(* IEC 61131-3 sources: daoli-st-library/_tools/rusty, 1 file *)

(* ---- iec_std_stub.st ---- *)
(* ============================================================================
   iec_std_stub.st  ——  道莅 L2 编译闸：IEC 61131-3 标准库外部声明桩
   ----------------------------------------------------------------------------
   用途：RuSTy (plc.exe) 不内建 IEC 标准函数/标准 FB 的声明，裸编译会把
        ABS/TON/R_TRIG 等判为 "Unknown type / Could not resolve reference"。
        本文件以 {external} 声明标准件接口，仅作 --check 夹具，不产生实现。

   纪律：
   1. 本文件**不属于**代码库交付物，只放在 _tools/rusty/ 下，不入 INDEX_REGISTRY。
   2. 声明按 IEC 61131-3 第 3 版标准语义书写，与各件源码零耦合。
   3. 泛型用 ANY_NUM / ANY_ELEMENTARY 表达，避免为每种位宽写重复声明。
   ============================================================================ *)

{external}
FUNCTION ABS<T: ANY_NUM> : T
VAR_INPUT IN : T; END_VAR
END_FUNCTION

{external}
FUNCTION SQRT<T: ANY_REAL> : T
VAR_INPUT IN : T; END_VAR
END_FUNCTION

{external}
FUNCTION LN<T: ANY_REAL> : T
VAR_INPUT IN : T; END_VAR
END_FUNCTION

{external}
FUNCTION LOG<T: ANY_REAL> : T
VAR_INPUT IN : T; END_VAR
END_FUNCTION

{external}
FUNCTION EXP<T: ANY_REAL> : T
VAR_INPUT IN : T; END_VAR
END_FUNCTION

{external}
FUNCTION SIN<T: ANY_REAL> : T
VAR_INPUT IN : T; END_VAR
END_FUNCTION

{external}
FUNCTION COS<T: ANY_REAL> : T
VAR_INPUT IN : T; END_VAR
END_FUNCTION

{external}
FUNCTION TAN<T: ANY_REAL> : T
VAR_INPUT IN : T; END_VAR
END_FUNCTION

{external}
FUNCTION ASIN<T: ANY_REAL> : T
VAR_INPUT IN : T; END_VAR
END_FUNCTION

{external}
FUNCTION ACOS<T: ANY_REAL> : T
VAR_INPUT IN : T; END_VAR
END_FUNCTION

{external}
FUNCTION ATAN<T: ANY_REAL> : T
VAR_INPUT IN : T; END_VAR
END_FUNCTION

{external}
FUNCTION EXPT<T: ANY_REAL> : T
VAR_INPUT IN1 : T; IN2 : T; END_VAR
END_FUNCTION

{external}
FUNCTION TRUNC<T: ANY_REAL> : T
VAR_INPUT IN : T; END_VAR
END_FUNCTION

{external}
FUNCTION ROUND<T: ANY_REAL> : T
VAR_INPUT IN : T; END_VAR
END_FUNCTION

{external}
FUNCTION FLOOR<T: ANY_REAL> : T
VAR_INPUT IN : T; END_VAR
END_FUNCTION

{external}
FUNCTION CEIL<T: ANY_REAL> : T
VAR_INPUT IN : T; END_VAR
END_FUNCTION

{external}
FUNCTION MIN<T: ANY_ELEMENTARY> : T
VAR_INPUT IN1 : T; IN2 : T; END_VAR
END_FUNCTION

{external}
FUNCTION MAX<T: ANY_ELEMENTARY> : T
VAR_INPUT IN1 : T; IN2 : T; END_VAR
END_FUNCTION

{external}
FUNCTION LIMIT<T: ANY_ELEMENTARY> : T
VAR_INPUT MN : T; IN : T; MX : T; END_VAR
END_FUNCTION

{external}
FUNCTION SEL<T: ANY_ELEMENTARY> : T
VAR_INPUT G : BOOL; IN0 : T; IN1 : T; END_VAR
END_FUNCTION

{external}
FUNCTION MUX<T: ANY_ELEMENTARY> : T
VAR_INPUT K : INT; IN0 : T; IN1 : T; IN2 : T; IN3 : T; END_VAR
END_FUNCTION

{external}
FUNCTION SHL<T: ANY_BIT> : T
VAR_INPUT IN : T; N : INT; END_VAR
END_FUNCTION

{external}
FUNCTION SHR<T: ANY_BIT> : T
VAR_INPUT IN : T; N : INT; END_VAR
END_FUNCTION

{external}
FUNCTION ROL<T: ANY_BIT> : T
VAR_INPUT IN : T; N : INT; END_VAR
END_FUNCTION

{external}
FUNCTION ROR<T: ANY_BIT> : T
VAR_INPUT IN : T; N : INT; END_VAR
END_FUNCTION

(* ---- 字符串九函数 ---- *)
{external}
FUNCTION LEN : UDINT
VAR_INPUT IN : STRING; END_VAR
END_FUNCTION

{external}
FUNCTION LEFT : STRING
VAR_INPUT IN : STRING; L : UDINT; END_VAR
END_FUNCTION

{external}
FUNCTION RIGHT : STRING
VAR_INPUT IN : STRING; L : UDINT; END_VAR
END_FUNCTION

{external}
FUNCTION MID : STRING
VAR_INPUT IN : STRING; L : UDINT; P : UDINT := 1; END_VAR
END_FUNCTION

{external}
FUNCTION CONCAT : STRING
VAR_INPUT IN1 : STRING; IN2 : STRING := ''; IN3 : STRING := ''; IN4 : STRING := ''; END_VAR
END_FUNCTION

{external}
FUNCTION INSERT : STRING
VAR_INPUT IN1 : STRING; IN2 : STRING; P : UDINT; END_VAR
END_FUNCTION

{external}
FUNCTION DELETE : STRING
VAR_INPUT IN : STRING; L : UDINT; P : UDINT; END_VAR
END_FUNCTION

{external}
FUNCTION REPLACE : STRING
VAR_INPUT IN1 : STRING; IN2 : STRING; L : UDINT; P : UDINT; END_VAR
END_FUNCTION

{external}
FUNCTION FIND : UDINT
VAR_INPUT IN1 : STRING; IN2 : STRING; END_VAR
END_FUNCTION

{external}
FUNCTION STRING_EQUAL : BOOL
VAR_INPUT a : STRING; b : STRING; END_VAR
END_FUNCTION

{external}
FUNCTION STRING_GREATER : BOOL
VAR_INPUT a : STRING; b : STRING; END_VAR
END_FUNCTION

{external}
FUNCTION STRING_LESS : BOOL
VAR_INPUT a : STRING; b : STRING; END_VAR
END_FUNCTION

{external}
FUNCTION WSTRING_EQUAL : BOOL
VAR_INPUT a : WSTRING; b : WSTRING; END_VAR
END_FUNCTION

(* ---- 标准边沿/定时/计数 FB（空体声明，仅满足类型解析） ---- *)
FUNCTION_BLOCK TON
VAR_INPUT
    IN : BOOL;
    PT : TIME;
END_VAR
VAR_OUTPUT
    Q : BOOL;
    ET : TIME;
END_VAR
END_FUNCTION_BLOCK

FUNCTION_BLOCK TOF
VAR_INPUT
    IN : BOOL;
    PT : TIME;
END_VAR
VAR_OUTPUT
    Q : BOOL;
    ET : TIME;
END_VAR
END_FUNCTION_BLOCK

FUNCTION_BLOCK TP
VAR_INPUT
    IN : BOOL;
    PT : TIME;
END_VAR
VAR_OUTPUT
    Q : BOOL;
    ET : TIME;
END_VAR
END_FUNCTION_BLOCK

FUNCTION_BLOCK R_TRIG
VAR_INPUT
    CLK : BOOL;
END_VAR
VAR_OUTPUT
    Q : BOOL;
END_VAR
END_FUNCTION_BLOCK

FUNCTION_BLOCK F_TRIG
VAR_INPUT
    CLK : BOOL;
END_VAR
VAR_OUTPUT
    Q : BOOL;
END_VAR
END_FUNCTION_BLOCK

FUNCTION_BLOCK CTU
VAR_INPUT
    CU : BOOL;
    R : BOOL;
    PV : INT;
END_VAR
VAR_OUTPUT
    Q : BOOL;
    CV : INT;
END_VAR
END_FUNCTION_BLOCK

FUNCTION_BLOCK CTD
VAR_INPUT
    CD : BOOL;
    LD : BOOL;
    PV : INT;
END_VAR
VAR_OUTPUT
    Q : BOOL;
    CV : INT;
END_VAR
END_FUNCTION_BLOCK

FUNCTION_BLOCK CTUD
VAR_INPUT
    CU : BOOL;
    CD : BOOL;
    R : BOOL;
    LD : BOOL;
    PV : INT;
END_VAR
VAR_OUTPUT
    QU : BOOL;
    QD : BOOL;
    CV : INT;
END_VAR
END_FUNCTION_BLOCK

(* ---- R71 补：类型转换 / ATAN2 / MOVE ---- *)
{external}
FUNCTION TIME_TO_REAL : REAL
VAR_INPUT IN : TIME; END_VAR
END_FUNCTION

{external}
FUNCTION TIME_TO_LREAL : LREAL
VAR_INPUT IN : TIME; END_VAR
END_FUNCTION

{external}
FUNCTION TIME_TO_DINT : DINT
VAR_INPUT IN : TIME; END_VAR
END_FUNCTION

{external}
FUNCTION TIME_TO_UDINT : UDINT
VAR_INPUT IN : TIME; END_VAR
END_FUNCTION

{external}
FUNCTION TIME_TO_LINT : LINT
VAR_INPUT IN : TIME; END_VAR
END_FUNCTION

{external}
FUNCTION UDINT_TO_REAL : REAL
VAR_INPUT IN : UDINT; END_VAR
END_FUNCTION

{external}
FUNCTION UDINT_TO_LREAL : LREAL
VAR_INPUT IN : UDINT; END_VAR
END_FUNCTION

{external}
FUNCTION UDINT_TO_DINT : DINT
VAR_INPUT IN : UDINT; END_VAR
END_FUNCTION

{external}
FUNCTION DINT_TO_REAL : REAL
VAR_INPUT IN : DINT; END_VAR
END_FUNCTION

{external}
FUNCTION DINT_TO_LREAL : LREAL
VAR_INPUT IN : DINT; END_VAR
END_FUNCTION

{external}
FUNCTION INT_TO_REAL : REAL
VAR_INPUT IN : INT; END_VAR
END_FUNCTION

{external}
FUNCTION INT_TO_LREAL : LREAL
VAR_INPUT IN : INT; END_VAR
END_FUNCTION

{external}
FUNCTION REAL_TO_DINT : DINT
VAR_INPUT IN : REAL; END_VAR
END_FUNCTION

{external}
FUNCTION REAL_TO_INT : INT
VAR_INPUT IN : REAL; END_VAR
END_FUNCTION

{external}
FUNCTION REAL_TO_UDINT : UDINT
VAR_INPUT IN : REAL; END_VAR
END_FUNCTION

{external}
FUNCTION LREAL_TO_REAL : REAL
VAR_INPUT IN : LREAL; END_VAR
END_FUNCTION

{external}
FUNCTION REAL_TO_LREAL : LREAL
VAR_INPUT IN : REAL; END_VAR
END_FUNCTION

{external}
FUNCTION LREAL_TO_DINT : DINT
VAR_INPUT IN : LREAL; END_VAR
END_FUNCTION

{external}
FUNCTION LREAL_TO_UDINT : UDINT
VAR_INPUT IN : LREAL; END_VAR
END_FUNCTION

{external}
FUNCTION BOOL_TO_INT : INT
VAR_INPUT IN : BOOL; END_VAR
END_FUNCTION

{external}
FUNCTION BOOL_TO_WORD : WORD
VAR_INPUT IN : BOOL; END_VAR
END_FUNCTION

{external}
FUNCTION WORD_TO_INT : INT
VAR_INPUT IN : WORD; END_VAR
END_FUNCTION

{external}
FUNCTION INT_TO_WORD : WORD
VAR_INPUT IN : INT; END_VAR
END_FUNCTION

{external}
FUNCTION WORD_TO_BOOL : BOOL
VAR_INPUT IN : WORD; END_VAR
END_FUNCTION

{external}
FUNCTION BYTE_TO_INT : INT
VAR_INPUT IN : BYTE; END_VAR
END_FUNCTION

{external}
FUNCTION INT_TO_BYTE : BYTE
VAR_INPUT IN : INT; END_VAR
END_FUNCTION

{external}
FUNCTION DT_TO_DINT : DINT
VAR_INPUT IN : DATE_AND_TIME; END_VAR
END_FUNCTION

{external}
FUNCTION DINT_TO_DT : DATE_AND_TIME
VAR_INPUT IN : DINT; END_VAR
END_FUNCTION

{external}
FUNCTION TOD_TO_DINT : DINT
VAR_INPUT IN : TIME_OF_DAY; END_VAR
END_FUNCTION

{external}
FUNCTION DINT_TO_TOD : TIME_OF_DAY
VAR_INPUT IN : DINT; END_VAR
END_FUNCTION

{external}
FUNCTION ATAN2<T: ANY_REAL> : T
VAR_INPUT Y : T; X : T; END_VAR
END_FUNCTION

{external}
FUNCTION MOVE<T: ANY_ELEMENTARY> : T
VAR_INPUT IN : T; END_VAR
END_FUNCTION

(* ---- R71 补二：时间域与位宽转换 ---- *)

{external}
FUNCTION DINT_TO_TIME : TIME
VAR_INPUT IN : DINT; END_VAR
END_FUNCTION

{external}
FUNCTION INT_TO_TIME : TIME
VAR_INPUT IN : INT; END_VAR
END_FUNCTION

{external}
FUNCTION UDINT_TO_TIME : TIME
VAR_INPUT IN : UDINT; END_VAR
END_FUNCTION

{external}
FUNCTION REAL_TO_TIME : TIME
VAR_INPUT IN : REAL; END_VAR
END_FUNCTION

{external}
FUNCTION LREAL_TO_TIME : TIME
VAR_INPUT IN : LREAL; END_VAR
END_FUNCTION

{external}
FUNCTION TIME_TO_INT : INT
VAR_INPUT IN : TIME; END_VAR
END_FUNCTION

{external}
FUNCTION DWORD_TO_DINT : DINT
VAR_INPUT IN : DWORD; END_VAR
END_FUNCTION

{external}
FUNCTION DINT_TO_DWORD : DWORD
VAR_INPUT IN : DINT; END_VAR
END_FUNCTION

{external}
FUNCTION LWORD_TO_LINT : LINT
VAR_INPUT IN : LWORD; END_VAR
END_FUNCTION

{external}
FUNCTION LINT_TO_LWORD : LWORD
VAR_INPUT IN : LINT; END_VAR
END_FUNCTION

{external}
FUNCTION WORD_TO_DWORD : DWORD
VAR_INPUT IN : WORD; END_VAR
END_FUNCTION

{external}
FUNCTION BYTE_TO_WORD : WORD
VAR_INPUT IN : BYTE; END_VAR
END_FUNCTION

{external}
FUNCTION TOD_TO_TIME : TIME
VAR_INPUT IN : TIME_OF_DAY; END_VAR
END_FUNCTION

{external}
FUNCTION TIME_TO_TOD : TIME_OF_DAY
VAR_INPUT IN : TIME; END_VAR
END_FUNCTION

(* ---- R71 补三：有/无符号与位宽互转 ---- *)

{external}
FUNCTION DINT_TO_UDINT : UDINT
VAR_INPUT IN : DINT; END_VAR
END_FUNCTION

{external}
FUNCTION UDINT_TO_INT : INT
VAR_INPUT IN : UDINT; END_VAR
END_FUNCTION

{external}
FUNCTION INT_TO_UDINT : UDINT
VAR_INPUT IN : INT; END_VAR
END_FUNCTION

{external}
FUNCTION LINT_TO_DINT : DINT
VAR_INPUT IN : LINT; END_VAR
END_FUNCTION

{external}
FUNCTION DINT_TO_LINT : LINT
VAR_INPUT IN : DINT; END_VAR
END_FUNCTION

{external}
FUNCTION WORD_TO_UDINT : UDINT
VAR_INPUT IN : WORD; END_VAR
END_FUNCTION

{external}
FUNCTION UDINT_TO_WORD : WORD
VAR_INPUT IN : UDINT; END_VAR
END_FUNCTION

{external}
FUNCTION BYTE_TO_UDINT : UDINT
VAR_INPUT IN : BYTE; END_VAR
END_FUNCTION

{external}
FUNCTION TIME_TO_WORD : WORD
VAR_INPUT IN : TIME; END_VAR
END_FUNCTION

(* ===== BEGIN AUTO-GENERATED CONVERSIONS  (stub_fix.py 维护，勿手改) ===== *)
(* 由 _tools/stub_fix.py 自动生成，覆盖全部 IEC 61131-3 标准转换。 *)

{external}
FUNCTION BYTE_TO_DINT : DINT
VAR_INPUT IN : BYTE; END_VAR
END_FUNCTION

{external}
FUNCTION BYTE_TO_DWORD : DWORD
VAR_INPUT IN : BYTE; END_VAR
END_FUNCTION

{external}
FUNCTION BYTE_TO_LINT : LINT
VAR_INPUT IN : BYTE; END_VAR
END_FUNCTION

{external}
FUNCTION BYTE_TO_LREAL : LREAL
VAR_INPUT IN : BYTE; END_VAR
END_FUNCTION

{external}
FUNCTION BYTE_TO_LWORD : LWORD
VAR_INPUT IN : BYTE; END_VAR
END_FUNCTION

{external}
FUNCTION BYTE_TO_REAL : REAL
VAR_INPUT IN : BYTE; END_VAR
END_FUNCTION

{external}
FUNCTION BYTE_TO_SINT : SINT
VAR_INPUT IN : BYTE; END_VAR
END_FUNCTION

{external}
FUNCTION BYTE_TO_STRING : STRING
VAR_INPUT IN : BYTE; END_VAR
END_FUNCTION

{external}
FUNCTION BYTE_TO_UINT : UINT
VAR_INPUT IN : BYTE; END_VAR
END_FUNCTION

{external}
FUNCTION BYTE_TO_ULINT : ULINT
VAR_INPUT IN : BYTE; END_VAR
END_FUNCTION

{external}
FUNCTION BYTE_TO_USINT : USINT
VAR_INPUT IN : BYTE; END_VAR
END_FUNCTION

{external}
FUNCTION DATE_TO_DINT : DINT
VAR_INPUT IN : DATE; END_VAR
END_FUNCTION

{external}
FUNCTION DATE_TO_DT : DT
VAR_INPUT IN : DATE; END_VAR
END_FUNCTION

{external}
FUNCTION DATE_TO_DTL : DTL
VAR_INPUT IN : DATE; END_VAR
END_FUNCTION

{external}
FUNCTION DATE_TO_INT : INT
VAR_INPUT IN : DATE; END_VAR
END_FUNCTION

{external}
FUNCTION DATE_TO_LINT : LINT
VAR_INPUT IN : DATE; END_VAR
END_FUNCTION

{external}
FUNCTION DATE_TO_LREAL : LREAL
VAR_INPUT IN : DATE; END_VAR
END_FUNCTION

{external}
FUNCTION DATE_TO_REAL : REAL
VAR_INPUT IN : DATE; END_VAR
END_FUNCTION

{external}
FUNCTION DATE_TO_STRING : STRING
VAR_INPUT IN : DATE; END_VAR
END_FUNCTION

{external}
FUNCTION DATE_TO_TIME : TIME
VAR_INPUT IN : DATE; END_VAR
END_FUNCTION

{external}
FUNCTION DATE_TO_TOD : TOD
VAR_INPUT IN : DATE; END_VAR
END_FUNCTION

{external}
FUNCTION DATE_TO_UDINT : UDINT
VAR_INPUT IN : DATE; END_VAR
END_FUNCTION

{external}
FUNCTION DINT_TO_BYTE : BYTE
VAR_INPUT IN : DINT; END_VAR
END_FUNCTION

{external}
FUNCTION DINT_TO_DATE : DATE
VAR_INPUT IN : DINT; END_VAR
END_FUNCTION

{external}
FUNCTION DINT_TO_INT : INT
VAR_INPUT IN : DINT; END_VAR
END_FUNCTION

{external}
FUNCTION DINT_TO_LWORD : LWORD
VAR_INPUT IN : DINT; END_VAR
END_FUNCTION

{external}
FUNCTION DINT_TO_SINT : SINT
VAR_INPUT IN : DINT; END_VAR
END_FUNCTION

{external}
FUNCTION DINT_TO_STRING : STRING
VAR_INPUT IN : DINT; END_VAR
END_FUNCTION

{external}
FUNCTION DINT_TO_UINT : UINT
VAR_INPUT IN : DINT; END_VAR
END_FUNCTION

{external}
FUNCTION DINT_TO_ULINT : ULINT
VAR_INPUT IN : DINT; END_VAR
END_FUNCTION

{external}
FUNCTION DINT_TO_USINT : USINT
VAR_INPUT IN : DINT; END_VAR
END_FUNCTION

{external}
FUNCTION DINT_TO_WORD : WORD
VAR_INPUT IN : DINT; END_VAR
END_FUNCTION

{external}
FUNCTION DTL_TO_DATE : DATE
VAR_INPUT IN : DTL; END_VAR
END_FUNCTION

{external}
FUNCTION DTL_TO_DINT : DINT
VAR_INPUT IN : DTL; END_VAR
END_FUNCTION

{external}
FUNCTION DTL_TO_DT : DT
VAR_INPUT IN : DTL; END_VAR
END_FUNCTION

{external}
FUNCTION DTL_TO_INT : INT
VAR_INPUT IN : DTL; END_VAR
END_FUNCTION

{external}
FUNCTION DTL_TO_LINT : LINT
VAR_INPUT IN : DTL; END_VAR
END_FUNCTION

{external}
FUNCTION DTL_TO_LREAL : LREAL
VAR_INPUT IN : DTL; END_VAR
END_FUNCTION

{external}
FUNCTION DTL_TO_REAL : REAL
VAR_INPUT IN : DTL; END_VAR
END_FUNCTION

{external}
FUNCTION DTL_TO_STRING : STRING
VAR_INPUT IN : DTL; END_VAR
END_FUNCTION

{external}
FUNCTION DTL_TO_TIME : TIME
VAR_INPUT IN : DTL; END_VAR
END_FUNCTION

{external}
FUNCTION DTL_TO_TOD : TOD
VAR_INPUT IN : DTL; END_VAR
END_FUNCTION

{external}
FUNCTION DTL_TO_UDINT : UDINT
VAR_INPUT IN : DTL; END_VAR
END_FUNCTION

{external}
FUNCTION DT_TO_DATE : DATE
VAR_INPUT IN : DT; END_VAR
END_FUNCTION

{external}
FUNCTION DT_TO_DTL : DTL
VAR_INPUT IN : DT; END_VAR
END_FUNCTION

{external}
FUNCTION DT_TO_INT : INT
VAR_INPUT IN : DT; END_VAR
END_FUNCTION

{external}
FUNCTION DT_TO_LINT : LINT
VAR_INPUT IN : DT; END_VAR
END_FUNCTION

{external}
FUNCTION DT_TO_LREAL : LREAL
VAR_INPUT IN : DT; END_VAR
END_FUNCTION

{external}
FUNCTION DT_TO_REAL : REAL
VAR_INPUT IN : DT; END_VAR
END_FUNCTION

{external}
FUNCTION DT_TO_STRING : STRING
VAR_INPUT IN : DT; END_VAR
END_FUNCTION

{external}
FUNCTION DT_TO_TIME : TIME
VAR_INPUT IN : DT; END_VAR
END_FUNCTION

{external}
FUNCTION DT_TO_TOD : TOD
VAR_INPUT IN : DT; END_VAR
END_FUNCTION

{external}
FUNCTION DT_TO_UDINT : UDINT
VAR_INPUT IN : DT; END_VAR
END_FUNCTION

{external}
FUNCTION DWORD_TO_BYTE : BYTE
VAR_INPUT IN : DWORD; END_VAR
END_FUNCTION

{external}
FUNCTION DWORD_TO_INT : INT
VAR_INPUT IN : DWORD; END_VAR
END_FUNCTION

{external}
FUNCTION DWORD_TO_LINT : LINT
VAR_INPUT IN : DWORD; END_VAR
END_FUNCTION

{external}
FUNCTION DWORD_TO_LREAL : LREAL
VAR_INPUT IN : DWORD; END_VAR
END_FUNCTION

{external}
FUNCTION DWORD_TO_LWORD : LWORD
VAR_INPUT IN : DWORD; END_VAR
END_FUNCTION

{external}
FUNCTION DWORD_TO_REAL : REAL
VAR_INPUT IN : DWORD; END_VAR
END_FUNCTION

{external}
FUNCTION DWORD_TO_SINT : SINT
VAR_INPUT IN : DWORD; END_VAR
END_FUNCTION

{external}
FUNCTION DWORD_TO_STRING : STRING
VAR_INPUT IN : DWORD; END_VAR
END_FUNCTION

{external}
FUNCTION DWORD_TO_UDINT : UDINT
VAR_INPUT IN : DWORD; END_VAR
END_FUNCTION

{external}
FUNCTION DWORD_TO_UINT : UINT
VAR_INPUT IN : DWORD; END_VAR
END_FUNCTION

{external}
FUNCTION DWORD_TO_ULINT : ULINT
VAR_INPUT IN : DWORD; END_VAR
END_FUNCTION

{external}
FUNCTION DWORD_TO_USINT : USINT
VAR_INPUT IN : DWORD; END_VAR
END_FUNCTION

{external}
FUNCTION DWORD_TO_WORD : WORD
VAR_INPUT IN : DWORD; END_VAR
END_FUNCTION

{external}
FUNCTION INT_TO_DATE : DATE
VAR_INPUT IN : INT; END_VAR
END_FUNCTION

{external}
FUNCTION INT_TO_DINT : DINT
VAR_INPUT IN : INT; END_VAR
END_FUNCTION

{external}
FUNCTION INT_TO_DT : DT
VAR_INPUT IN : INT; END_VAR
END_FUNCTION

{external}
FUNCTION INT_TO_DWORD : DWORD
VAR_INPUT IN : INT; END_VAR
END_FUNCTION

{external}
FUNCTION INT_TO_LINT : LINT
VAR_INPUT IN : INT; END_VAR
END_FUNCTION

{external}
FUNCTION INT_TO_LWORD : LWORD
VAR_INPUT IN : INT; END_VAR
END_FUNCTION

{external}
FUNCTION INT_TO_SINT : SINT
VAR_INPUT IN : INT; END_VAR
END_FUNCTION

{external}
FUNCTION INT_TO_STRING : STRING
VAR_INPUT IN : INT; END_VAR
END_FUNCTION

{external}
FUNCTION INT_TO_TOD : TOD
VAR_INPUT IN : INT; END_VAR
END_FUNCTION

{external}
FUNCTION INT_TO_UINT : UINT
VAR_INPUT IN : INT; END_VAR
END_FUNCTION

{external}
FUNCTION INT_TO_ULINT : ULINT
VAR_INPUT IN : INT; END_VAR
END_FUNCTION

{external}
FUNCTION INT_TO_USINT : USINT
VAR_INPUT IN : INT; END_VAR
END_FUNCTION

{external}
FUNCTION LINT_TO_BYTE : BYTE
VAR_INPUT IN : LINT; END_VAR
END_FUNCTION

{external}
FUNCTION LINT_TO_DATE : DATE
VAR_INPUT IN : LINT; END_VAR
END_FUNCTION

{external}
FUNCTION LINT_TO_DT : DT
VAR_INPUT IN : LINT; END_VAR
END_FUNCTION

{external}
FUNCTION LINT_TO_DWORD : DWORD
VAR_INPUT IN : LINT; END_VAR
END_FUNCTION

{external}
FUNCTION LINT_TO_INT : INT
VAR_INPUT IN : LINT; END_VAR
END_FUNCTION

{external}
FUNCTION LINT_TO_LREAL : LREAL
VAR_INPUT IN : LINT; END_VAR
END_FUNCTION

{external}
FUNCTION LINT_TO_REAL : REAL
VAR_INPUT IN : LINT; END_VAR
END_FUNCTION

{external}
FUNCTION LINT_TO_SINT : SINT
VAR_INPUT IN : LINT; END_VAR
END_FUNCTION

{external}
FUNCTION LINT_TO_STRING : STRING
VAR_INPUT IN : LINT; END_VAR
END_FUNCTION

{external}
FUNCTION LINT_TO_TIME : TIME
VAR_INPUT IN : LINT; END_VAR
END_FUNCTION

{external}
FUNCTION LINT_TO_TOD : TOD
VAR_INPUT IN : LINT; END_VAR
END_FUNCTION

{external}
FUNCTION LINT_TO_UDINT : UDINT
VAR_INPUT IN : LINT; END_VAR
END_FUNCTION

{external}
FUNCTION LINT_TO_UINT : UINT
VAR_INPUT IN : LINT; END_VAR
END_FUNCTION

{external}
FUNCTION LINT_TO_ULINT : ULINT
VAR_INPUT IN : LINT; END_VAR
END_FUNCTION

{external}
FUNCTION LINT_TO_USINT : USINT
VAR_INPUT IN : LINT; END_VAR
END_FUNCTION

{external}
FUNCTION LINT_TO_WORD : WORD
VAR_INPUT IN : LINT; END_VAR
END_FUNCTION

{external}
FUNCTION LREAL_TO_BYTE : BYTE
VAR_INPUT IN : LREAL; END_VAR
END_FUNCTION

{external}
FUNCTION LREAL_TO_DATE : DATE
VAR_INPUT IN : LREAL; END_VAR
END_FUNCTION

{external}
FUNCTION LREAL_TO_DT : DT
VAR_INPUT IN : LREAL; END_VAR
END_FUNCTION

{external}
FUNCTION LREAL_TO_DWORD : DWORD
VAR_INPUT IN : LREAL; END_VAR
END_FUNCTION

{external}
FUNCTION LREAL_TO_INT : INT
VAR_INPUT IN : LREAL; END_VAR
END_FUNCTION

{external}
FUNCTION LREAL_TO_LINT : LINT
VAR_INPUT IN : LREAL; END_VAR
END_FUNCTION

{external}
FUNCTION LREAL_TO_LWORD : LWORD
VAR_INPUT IN : LREAL; END_VAR
END_FUNCTION

{external}
FUNCTION LREAL_TO_SINT : SINT
VAR_INPUT IN : LREAL; END_VAR
END_FUNCTION

{external}
FUNCTION LREAL_TO_STRING : STRING
VAR_INPUT IN : LREAL; END_VAR
END_FUNCTION

{external}
FUNCTION LREAL_TO_TOD : TOD
VAR_INPUT IN : LREAL; END_VAR
END_FUNCTION

{external}
FUNCTION LREAL_TO_UINT : UINT
VAR_INPUT IN : LREAL; END_VAR
END_FUNCTION

{external}
FUNCTION LREAL_TO_ULINT : ULINT
VAR_INPUT IN : LREAL; END_VAR
END_FUNCTION

{external}
FUNCTION LREAL_TO_USINT : USINT
VAR_INPUT IN : LREAL; END_VAR
END_FUNCTION

{external}
FUNCTION LREAL_TO_WORD : WORD
VAR_INPUT IN : LREAL; END_VAR
END_FUNCTION

{external}
FUNCTION LWORD_TO_BYTE : BYTE
VAR_INPUT IN : LWORD; END_VAR
END_FUNCTION

{external}
FUNCTION LWORD_TO_DINT : DINT
VAR_INPUT IN : LWORD; END_VAR
END_FUNCTION

{external}
FUNCTION LWORD_TO_DWORD : DWORD
VAR_INPUT IN : LWORD; END_VAR
END_FUNCTION

{external}
FUNCTION LWORD_TO_INT : INT
VAR_INPUT IN : LWORD; END_VAR
END_FUNCTION

{external}
FUNCTION LWORD_TO_LREAL : LREAL
VAR_INPUT IN : LWORD; END_VAR
END_FUNCTION

{external}
FUNCTION LWORD_TO_REAL : REAL
VAR_INPUT IN : LWORD; END_VAR
END_FUNCTION

{external}
FUNCTION LWORD_TO_SINT : SINT
VAR_INPUT IN : LWORD; END_VAR
END_FUNCTION

{external}
FUNCTION LWORD_TO_STRING : STRING
VAR_INPUT IN : LWORD; END_VAR
END_FUNCTION

{external}
FUNCTION LWORD_TO_UDINT : UDINT
VAR_INPUT IN : LWORD; END_VAR
END_FUNCTION

{external}
FUNCTION LWORD_TO_UINT : UINT
VAR_INPUT IN : LWORD; END_VAR
END_FUNCTION

{external}
FUNCTION LWORD_TO_ULINT : ULINT
VAR_INPUT IN : LWORD; END_VAR
END_FUNCTION

{external}
FUNCTION LWORD_TO_USINT : USINT
VAR_INPUT IN : LWORD; END_VAR
END_FUNCTION

{external}
FUNCTION LWORD_TO_WORD : WORD
VAR_INPUT IN : LWORD; END_VAR
END_FUNCTION

{external}
FUNCTION REAL_TO_BYTE : BYTE
VAR_INPUT IN : REAL; END_VAR
END_FUNCTION

{external}
FUNCTION REAL_TO_DATE : DATE
VAR_INPUT IN : REAL; END_VAR
END_FUNCTION

{external}
FUNCTION REAL_TO_DT : DT
VAR_INPUT IN : REAL; END_VAR
END_FUNCTION

{external}
FUNCTION REAL_TO_DWORD : DWORD
VAR_INPUT IN : REAL; END_VAR
END_FUNCTION

{external}
FUNCTION REAL_TO_LINT : LINT
VAR_INPUT IN : REAL; END_VAR
END_FUNCTION

{external}
FUNCTION REAL_TO_LWORD : LWORD
VAR_INPUT IN : REAL; END_VAR
END_FUNCTION

{external}
FUNCTION REAL_TO_SINT : SINT
VAR_INPUT IN : REAL; END_VAR
END_FUNCTION

{external}
FUNCTION REAL_TO_STRING : STRING
VAR_INPUT IN : REAL; END_VAR
END_FUNCTION

{external}
FUNCTION REAL_TO_TOD : TOD
VAR_INPUT IN : REAL; END_VAR
END_FUNCTION

{external}
FUNCTION REAL_TO_UINT : UINT
VAR_INPUT IN : REAL; END_VAR
END_FUNCTION

{external}
FUNCTION REAL_TO_ULINT : ULINT
VAR_INPUT IN : REAL; END_VAR
END_FUNCTION

{external}
FUNCTION REAL_TO_USINT : USINT
VAR_INPUT IN : REAL; END_VAR
END_FUNCTION

{external}
FUNCTION REAL_TO_WORD : WORD
VAR_INPUT IN : REAL; END_VAR
END_FUNCTION

{external}
FUNCTION SINT_TO_BYTE : BYTE
VAR_INPUT IN : SINT; END_VAR
END_FUNCTION

{external}
FUNCTION SINT_TO_DINT : DINT
VAR_INPUT IN : SINT; END_VAR
END_FUNCTION

{external}
FUNCTION SINT_TO_DWORD : DWORD
VAR_INPUT IN : SINT; END_VAR
END_FUNCTION

{external}
FUNCTION SINT_TO_INT : INT
VAR_INPUT IN : SINT; END_VAR
END_FUNCTION

{external}
FUNCTION SINT_TO_LINT : LINT
VAR_INPUT IN : SINT; END_VAR
END_FUNCTION

{external}
FUNCTION SINT_TO_LREAL : LREAL
VAR_INPUT IN : SINT; END_VAR
END_FUNCTION

{external}
FUNCTION SINT_TO_LWORD : LWORD
VAR_INPUT IN : SINT; END_VAR
END_FUNCTION

{external}
FUNCTION SINT_TO_REAL : REAL
VAR_INPUT IN : SINT; END_VAR
END_FUNCTION

{external}
FUNCTION SINT_TO_STRING : STRING
VAR_INPUT IN : SINT; END_VAR
END_FUNCTION

{external}
FUNCTION SINT_TO_UDINT : UDINT
VAR_INPUT IN : SINT; END_VAR
END_FUNCTION

{external}
FUNCTION SINT_TO_UINT : UINT
VAR_INPUT IN : SINT; END_VAR
END_FUNCTION

{external}
FUNCTION SINT_TO_ULINT : ULINT
VAR_INPUT IN : SINT; END_VAR
END_FUNCTION

{external}
FUNCTION SINT_TO_USINT : USINT
VAR_INPUT IN : SINT; END_VAR
END_FUNCTION

{external}
FUNCTION SINT_TO_WORD : WORD
VAR_INPUT IN : SINT; END_VAR
END_FUNCTION

{external}
FUNCTION STRING_TO_BYTE : BYTE
VAR_INPUT IN : STRING; END_VAR
END_FUNCTION

{external}
FUNCTION STRING_TO_DATE : DATE
VAR_INPUT IN : STRING; END_VAR
END_FUNCTION

{external}
FUNCTION STRING_TO_DINT : DINT
VAR_INPUT IN : STRING; END_VAR
END_FUNCTION

{external}
FUNCTION STRING_TO_DT : DT
VAR_INPUT IN : STRING; END_VAR
END_FUNCTION

{external}
FUNCTION STRING_TO_DTL : DTL
VAR_INPUT IN : STRING; END_VAR
END_FUNCTION

{external}
FUNCTION STRING_TO_DWORD : DWORD
VAR_INPUT IN : STRING; END_VAR
END_FUNCTION

{external}
FUNCTION STRING_TO_INT : INT
VAR_INPUT IN : STRING; END_VAR
END_FUNCTION

{external}
FUNCTION STRING_TO_LINT : LINT
VAR_INPUT IN : STRING; END_VAR
END_FUNCTION

{external}
FUNCTION STRING_TO_LREAL : LREAL
VAR_INPUT IN : STRING; END_VAR
END_FUNCTION

{external}
FUNCTION STRING_TO_LWORD : LWORD
VAR_INPUT IN : STRING; END_VAR
END_FUNCTION

{external}
FUNCTION STRING_TO_REAL : REAL
VAR_INPUT IN : STRING; END_VAR
END_FUNCTION

{external}
FUNCTION STRING_TO_SINT : SINT
VAR_INPUT IN : STRING; END_VAR
END_FUNCTION

{external}
FUNCTION STRING_TO_TIME : TIME
VAR_INPUT IN : STRING; END_VAR
END_FUNCTION

{external}
FUNCTION STRING_TO_TOD : TOD
VAR_INPUT IN : STRING; END_VAR
END_FUNCTION

{external}
FUNCTION STRING_TO_UDINT : UDINT
VAR_INPUT IN : STRING; END_VAR
END_FUNCTION

{external}
FUNCTION STRING_TO_UINT : UINT
VAR_INPUT IN : STRING; END_VAR
END_FUNCTION

{external}
FUNCTION STRING_TO_ULINT : ULINT
VAR_INPUT IN : STRING; END_VAR
END_FUNCTION

{external}
FUNCTION STRING_TO_USINT : USINT
VAR_INPUT IN : STRING; END_VAR
END_FUNCTION

{external}
FUNCTION STRING_TO_WORD : WORD
VAR_INPUT IN : STRING; END_VAR
END_FUNCTION

{external}
FUNCTION TIME_TO_DATE : DATE
VAR_INPUT IN : TIME; END_VAR
END_FUNCTION

{external}
FUNCTION TIME_TO_DT : DT
VAR_INPUT IN : TIME; END_VAR
END_FUNCTION

{external}
FUNCTION TIME_TO_DTL : DTL
VAR_INPUT IN : TIME; END_VAR
END_FUNCTION

{external}
FUNCTION TIME_TO_STRING : STRING
VAR_INPUT IN : TIME; END_VAR
END_FUNCTION

{external}
FUNCTION TOD_TO_DATE : DATE
VAR_INPUT IN : TOD; END_VAR
END_FUNCTION

{external}
FUNCTION TOD_TO_DT : DT
VAR_INPUT IN : TOD; END_VAR
END_FUNCTION

{external}
FUNCTION TOD_TO_DTL : DTL
VAR_INPUT IN : TOD; END_VAR
END_FUNCTION

{external}
FUNCTION TOD_TO_INT : INT
VAR_INPUT IN : TOD; END_VAR
END_FUNCTION

{external}
FUNCTION TOD_TO_LINT : LINT
VAR_INPUT IN : TOD; END_VAR
END_FUNCTION

{external}
FUNCTION TOD_TO_LREAL : LREAL
VAR_INPUT IN : TOD; END_VAR
END_FUNCTION

{external}
FUNCTION TOD_TO_REAL : REAL
VAR_INPUT IN : TOD; END_VAR
END_FUNCTION

{external}
FUNCTION TOD_TO_STRING : STRING
VAR_INPUT IN : TOD; END_VAR
END_FUNCTION

{external}
FUNCTION TOD_TO_UDINT : UDINT
VAR_INPUT IN : TOD; END_VAR
END_FUNCTION

{external}
FUNCTION UDINT_TO_BYTE : BYTE
VAR_INPUT IN : UDINT; END_VAR
END_FUNCTION

{external}
FUNCTION UDINT_TO_DATE : DATE
VAR_INPUT IN : UDINT; END_VAR
END_FUNCTION

{external}
FUNCTION UDINT_TO_DT : DT
VAR_INPUT IN : UDINT; END_VAR
END_FUNCTION

{external}
FUNCTION UDINT_TO_DWORD : DWORD
VAR_INPUT IN : UDINT; END_VAR
END_FUNCTION

{external}
FUNCTION UDINT_TO_LINT : LINT
VAR_INPUT IN : UDINT; END_VAR
END_FUNCTION

{external}
FUNCTION UDINT_TO_LWORD : LWORD
VAR_INPUT IN : UDINT; END_VAR
END_FUNCTION

{external}
FUNCTION UDINT_TO_SINT : SINT
VAR_INPUT IN : UDINT; END_VAR
END_FUNCTION

{external}
FUNCTION UDINT_TO_STRING : STRING
VAR_INPUT IN : UDINT; END_VAR
END_FUNCTION

{external}
FUNCTION UDINT_TO_TOD : TOD
VAR_INPUT IN : UDINT; END_VAR
END_FUNCTION

{external}
FUNCTION UDINT_TO_UINT : UINT
VAR_INPUT IN : UDINT; END_VAR
END_FUNCTION

{external}
FUNCTION UDINT_TO_ULINT : ULINT
VAR_INPUT IN : UDINT; END_VAR
END_FUNCTION

{external}
FUNCTION UDINT_TO_USINT : USINT
VAR_INPUT IN : UDINT; END_VAR
END_FUNCTION

{external}
FUNCTION UINT_TO_BYTE : BYTE
VAR_INPUT IN : UINT; END_VAR
END_FUNCTION

{external}
FUNCTION UINT_TO_DINT : DINT
VAR_INPUT IN : UINT; END_VAR
END_FUNCTION

{external}
FUNCTION UINT_TO_DWORD : DWORD
VAR_INPUT IN : UINT; END_VAR
END_FUNCTION

{external}
FUNCTION UINT_TO_INT : INT
VAR_INPUT IN : UINT; END_VAR
END_FUNCTION

{external}
FUNCTION UINT_TO_LINT : LINT
VAR_INPUT IN : UINT; END_VAR
END_FUNCTION

{external}
FUNCTION UINT_TO_LREAL : LREAL
VAR_INPUT IN : UINT; END_VAR
END_FUNCTION

{external}
FUNCTION UINT_TO_LWORD : LWORD
VAR_INPUT IN : UINT; END_VAR
END_FUNCTION

{external}
FUNCTION UINT_TO_REAL : REAL
VAR_INPUT IN : UINT; END_VAR
END_FUNCTION

{external}
FUNCTION UINT_TO_SINT : SINT
VAR_INPUT IN : UINT; END_VAR
END_FUNCTION

{external}
FUNCTION UINT_TO_STRING : STRING
VAR_INPUT IN : UINT; END_VAR
END_FUNCTION

{external}
FUNCTION UINT_TO_UDINT : UDINT
VAR_INPUT IN : UINT; END_VAR
END_FUNCTION

{external}
FUNCTION UINT_TO_ULINT : ULINT
VAR_INPUT IN : UINT; END_VAR
END_FUNCTION

{external}
FUNCTION UINT_TO_USINT : USINT
VAR_INPUT IN : UINT; END_VAR
END_FUNCTION

{external}
FUNCTION UINT_TO_WORD : WORD
VAR_INPUT IN : UINT; END_VAR
END_FUNCTION

{external}
FUNCTION ULINT_TO_BYTE : BYTE
VAR_INPUT IN : ULINT; END_VAR
END_FUNCTION

{external}
FUNCTION ULINT_TO_DINT : DINT
VAR_INPUT IN : ULINT; END_VAR
END_FUNCTION

{external}
FUNCTION ULINT_TO_DWORD : DWORD
VAR_INPUT IN : ULINT; END_VAR
END_FUNCTION

{external}
FUNCTION ULINT_TO_INT : INT
VAR_INPUT IN : ULINT; END_VAR
END_FUNCTION

{external}
FUNCTION ULINT_TO_LINT : LINT
VAR_INPUT IN : ULINT; END_VAR
END_FUNCTION

{external}
FUNCTION ULINT_TO_LREAL : LREAL
VAR_INPUT IN : ULINT; END_VAR
END_FUNCTION

{external}
FUNCTION ULINT_TO_LWORD : LWORD
VAR_INPUT IN : ULINT; END_VAR
END_FUNCTION

{external}
FUNCTION ULINT_TO_REAL : REAL
VAR_INPUT IN : ULINT; END_VAR
END_FUNCTION

{external}
FUNCTION ULINT_TO_SINT : SINT
VAR_INPUT IN : ULINT; END_VAR
END_FUNCTION

{external}
FUNCTION ULINT_TO_STRING : STRING
VAR_INPUT IN : ULINT; END_VAR
END_FUNCTION

{external}
FUNCTION ULINT_TO_UDINT : UDINT
VAR_INPUT IN : ULINT; END_VAR
END_FUNCTION

{external}
FUNCTION ULINT_TO_UINT : UINT
VAR_INPUT IN : ULINT; END_VAR
END_FUNCTION

{external}
FUNCTION ULINT_TO_USINT : USINT
VAR_INPUT IN : ULINT; END_VAR
END_FUNCTION

{external}
FUNCTION ULINT_TO_WORD : WORD
VAR_INPUT IN : ULINT; END_VAR
END_FUNCTION

{external}
FUNCTION USINT_TO_BYTE : BYTE
VAR_INPUT IN : USINT; END_VAR
END_FUNCTION

{external}
FUNCTION USINT_TO_DINT : DINT
VAR_INPUT IN : USINT; END_VAR
END_FUNCTION

{external}
FUNCTION USINT_TO_DWORD : DWORD
VAR_INPUT IN : USINT; END_VAR
END_FUNCTION

{external}
FUNCTION USINT_TO_INT : INT
VAR_INPUT IN : USINT; END_VAR
END_FUNCTION

{external}
FUNCTION USINT_TO_LINT : LINT
VAR_INPUT IN : USINT; END_VAR
END_FUNCTION

{external}
FUNCTION USINT_TO_LREAL : LREAL
VAR_INPUT IN : USINT; END_VAR
END_FUNCTION

{external}
FUNCTION USINT_TO_LWORD : LWORD
VAR_INPUT IN : USINT; END_VAR
END_FUNCTION

{external}
FUNCTION USINT_TO_REAL : REAL
VAR_INPUT IN : USINT; END_VAR
END_FUNCTION

{external}
FUNCTION USINT_TO_SINT : SINT
VAR_INPUT IN : USINT; END_VAR
END_FUNCTION

{external}
FUNCTION USINT_TO_STRING : STRING
VAR_INPUT IN : USINT; END_VAR
END_FUNCTION

{external}
FUNCTION USINT_TO_UDINT : UDINT
VAR_INPUT IN : USINT; END_VAR
END_FUNCTION

{external}
FUNCTION USINT_TO_UINT : UINT
VAR_INPUT IN : USINT; END_VAR
END_FUNCTION

{external}
FUNCTION USINT_TO_ULINT : ULINT
VAR_INPUT IN : USINT; END_VAR
END_FUNCTION

{external}
FUNCTION USINT_TO_WORD : WORD
VAR_INPUT IN : USINT; END_VAR
END_FUNCTION

{external}
FUNCTION WORD_TO_BYTE : BYTE
VAR_INPUT IN : WORD; END_VAR
END_FUNCTION

{external}
FUNCTION WORD_TO_DINT : DINT
VAR_INPUT IN : WORD; END_VAR
END_FUNCTION

{external}
FUNCTION WORD_TO_LINT : LINT
VAR_INPUT IN : WORD; END_VAR
END_FUNCTION

{external}
FUNCTION WORD_TO_LREAL : LREAL
VAR_INPUT IN : WORD; END_VAR
END_FUNCTION

{external}
FUNCTION WORD_TO_LWORD : LWORD
VAR_INPUT IN : WORD; END_VAR
END_FUNCTION

{external}
FUNCTION WORD_TO_REAL : REAL
VAR_INPUT IN : WORD; END_VAR
END_FUNCTION

{external}
FUNCTION WORD_TO_SINT : SINT
VAR_INPUT IN : WORD; END_VAR
END_FUNCTION

{external}
FUNCTION WORD_TO_STRING : STRING
VAR_INPUT IN : WORD; END_VAR
END_FUNCTION

{external}
FUNCTION WORD_TO_UINT : UINT
VAR_INPUT IN : WORD; END_VAR
END_FUNCTION

{external}
FUNCTION WORD_TO_ULINT : ULINT
VAR_INPUT IN : WORD; END_VAR
END_FUNCTION

{external}
FUNCTION WORD_TO_USINT : USINT
VAR_INPUT IN : WORD; END_VAR
END_FUNCTION

(* ===== END AUTO-GENERATED CONVERSIONS ===== *)
